{attribute 'no_assign'}
{attribute 'call_after_init'}
FUNCTION_BLOCK FB_IED_WTURBINE EXTENDS FB_AcsiCommonIntelligentElectronicDeviceClass
VAR_INPUT
	WTURBINELD0: FB_LD_WTURBINELD0 := (bLinkResult:=THIS^.AddLogicalDeviceToContainer(ipLogicalDevice:=WTURBINELD0));
END_VAR
VAR
END_VAR

END_FUNCTION_BLOCK

(* stored: Version 1.1.0.1
   POU FB_IED_WTURBINE: Id {800a32bd-c2a8-4ee4-a3fd-60f721a9d4f0}, SpecialFunc None *)
